FUNCTION_BLOCK DebounceBool (* Migrated from IEC 61131-3 ST *)
  (* Standard: 61499-2 *)
  (* Version 1.0, 2026-11-06, st2fb *)
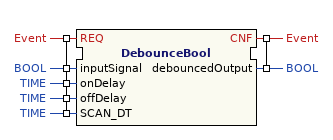
  EVENT_INPUT
    REQ WITH inputSignal, onDelay, offDelay, SCAN_DT;
  END_EVENT
  EVENT_OUTPUT
    CNF WITH debouncedOutput;
  END_EVENT
  VAR_INPUT
    inputSignal : BOOL;
    onDelay : TIME;
    offDelay : TIME;
    SCAN_DT : TIME;
  END_VAR
  VAR_OUTPUT
    debouncedOutput : BOOL;
  END_VAR
  VAR
    ST2FB_NOW : TIME := T#0s;
    tonTimer_IN : BOOL := FALSE;
    tonTimer_PT : TIME := T#0s;
    tonTimer_Q : BOOL := FALSE;
    tonTimer_ET : TIME := T#0s;
    tonTimer_STATE : INT := 0;
    tonTimer_PREV_IN : BOOL := FALSE;
    tonTimer_START_TIME : TIME := T#0s;
    tofTimer_IN : BOOL := FALSE;
    tofTimer_PT : TIME := T#0s;
    tofTimer_Q : BOOL := FALSE;
    tofTimer_ET : TIME := T#0s;
    tofTimer_STATE : INT := 0;
    tofTimer_PREV_IN : BOOL := FALSE;
    tofTimer_START_TIME : TIME := T#0s;
  END_VAR
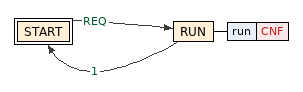
  EC_STATES
    START;
    RUN : run -> CNF;
  END_STATES
  EC_TRANSITIONS
    START TO RUN := REQ;
    RUN TO START := 1;
  END_TRANSITIONS
  ALGORITHM run IN ST:
ST2FB_NOW := ST2FB_NOW + SCAN_DT;

tonTimer_IN := inputSignal AND NOT debouncedOutput;
tonTimer_PT := onDelay;
IF (tonTimer_STATE = 0) AND NOT tonTimer_PREV_IN AND tonTimer_IN THEN
  tonTimer_STATE := 1;
  tonTimer_Q := FALSE;
  tonTimer_START_TIME := ST2FB_NOW;
ELSE
  IF NOT tonTimer_IN THEN
    tonTimer_ET := T#0s;
    tonTimer_Q := FALSE;
    tonTimer_STATE := 0;
  ELSIF tonTimer_STATE = 1 THEN
    IF tonTimer_START_TIME + tonTimer_PT <= ST2FB_NOW THEN
      tonTimer_STATE := 2;
      tonTimer_Q := TRUE;
      tonTimer_ET := tonTimer_PT;
    ELSE
      tonTimer_ET := ST2FB_NOW - tonTimer_START_TIME;
    END_IF;
  END_IF;
END_IF;
tonTimer_PREV_IN := tonTimer_IN;

tofTimer_IN := NOT inputSignal AND debouncedOutput;
tofTimer_PT := offDelay;
IF (tofTimer_STATE = 0) AND NOT tofTimer_PREV_IN AND tofTimer_IN THEN
  tofTimer_STATE := 1;
  tofTimer_Q := FALSE;
  tofTimer_START_TIME := ST2FB_NOW;
ELSE
  IF NOT tofTimer_IN THEN
    tofTimer_ET := T#0s;
    tofTimer_Q := FALSE;
    tofTimer_STATE := 0;
  ELSIF tofTimer_STATE = 1 THEN
    IF tofTimer_START_TIME + tofTimer_PT <= ST2FB_NOW THEN
      tofTimer_STATE := 2;
      tofTimer_Q := TRUE;
      tofTimer_ET := tofTimer_PT;
    ELSE
      tofTimer_ET := ST2FB_NOW - tofTimer_START_TIME;
    END_IF;
  END_IF;
END_IF;
tofTimer_PREV_IN := tofTimer_IN;

IF tonTimer_IN AND tonTimer_Q THEN
  debouncedOutput := TRUE;
ELSIF tofTimer_IN AND tofTimer_Q THEN
  debouncedOutput := FALSE;
END_IF;
  END_ALGORITHM
END_FUNCTION_BLOCK
